// TIA Portal V19 export
// export: Created 2026-10-15T09:44:23.7628945Z, ExportSetting WithDefaults, DisplayName Totally Integrated Automation Portal, DisplayVersion V19, DisplayName TIA Portal Openness, DisplayVersion V19, DisplayName TIA Portal Version Control Interface, DisplayVersion V19, DisplayName STEP 7 Professional, DisplayVersion V19, DisplayName STEP 7 Safety, DisplayVersion V19, DisplayName WinCC Basic/Comfort/Advanced, DisplayVersion V19, DisplayName WinCC Unified, DisplayVersion V19
FUNCTION "ROLL_PB9" : Void   // FC19, SCL
{ S7_Optimized_Access := 'TRUE' }
VERSION : 0.1
// stored: AutoNumber true, IsIECCheckEnabled false, SetENOAutomatically false, UDAEnableTagReadback false
   VAR_TEMP
      r : Bool;
      a1 : Word;
      a2 : Word;
      activeDataBlock : Int;
      comparisonResults : Array[0..0] of Bool;
   END_VAR
BEGIN

   #r := FALSE;
   #a1 := W#16#0000;
   #a2 := W#16#0000;
   #activeDataBlock := 0;
   // PB9, STEP 5 network 1
   #r := ((NOT "ROLL_State".M[32, 1]) AND (NOT "ROLL_State".M[32, 2]) AND "ROLL_IO".Input[0, 2]);
   "ROLL_State".M[32, 0] := #r;
   // PB9, STEP 5 network 2
   #r := "ROLL_State".M[32, 0];
   IF #r THEN
       "ROLL_State".M[32, 1] := TRUE;
   END_IF;
   #r := ((NOT "ROLL_IO".Input[0, 2]) OR "ROLL_IO".Input[0, 1] OR "ROLL_State".M[32, 2]);
   IF #r THEN
       "ROLL_State".M[32, 1] := FALSE;
   END_IF;
   // PB9, STEP 5 network 3
   #r := ((NOT "ROLL_IO".Input[0, 2]) OR "ROLL_IO".Input[0, 1]);
   "ROLL_State".M[32, 2] := #r;
   // PB9, STEP 5 network 4
   #r := ((NOT "ROLL_State".M[12, 0]) AND (NOT "ROLL_State".M[5, 0]) AND (NOT "ROLL_State".M[5, 2]) AND (NOT "ROLL_State".M[9, 0]));
   "ROLL_State".M[35, 1] := #r;
   // PB9, STEP 5 network 5
   #r := "ROLL_IO".Input[0, 4];
   IF #r THEN
       "ROLL_State".M[35, 2] := TRUE;
   END_IF;
   #r := ((NOT "ROLL_State".M[29, 0]) OR (NOT "ROLL_State".M[31, 5]) OR (NOT "ROLL_State".M[35, 1]) OR "ROLL_State".M[16, 3]);
   IF #r THEN
       "ROLL_State".M[35, 2] := FALSE;
   END_IF;
   // PB9, STEP 5 network 6
   #r := ("ROLL_State".M[32, 0] OR "ROLL_State".M[53, 6]);
   IF #r THEN
       "ROLL_State".M[37, 0] := TRUE;
   END_IF;
   #r := ("ROLL_State".M[32, 2] OR "ROLL_State".M[37, 1] OR "ROLL_State".M[38, 0] OR "ROLL_State".M[39, 5]);
   IF #r THEN
       "ROLL_State".M[37, 0] := FALSE;
   END_IF;
   // PB9, STEP 5 network 7
   #r := ((NOT "ROLL_IO".Input[123, 5]) AND (NOT "ROLL_IO".Input[123, 6]) AND (NOT "ROLL_State".M[53, 6]) AND "ROLL_State".M[31, 5] AND "ROLL_State".M[35, 2] AND "ROLL_State".M[37, 0]);
   IF #r THEN
       "ROLL_State".M[37, 1] := TRUE;
   END_IF;
   #r := ("ROLL_State".M[32, 2] OR "ROLL_State".M[37, 2] OR "ROLL_State".M[39, 6]);
   IF #r THEN
       "ROLL_State".M[37, 1] := FALSE;
   END_IF;
   // PB9, STEP 5 network 8
   #r := ((NOT "ROLL_IO".Output[113, 3]) AND (NOT "ROLL_State".M[9, 1]) AND (("ROLL_IO".Input[0, 5] AND "ROLL_IO".Input[14, 3] AND "ROLL_State".M[0, 4]) OR ("ROLL_IO".Input[123, 4] AND "ROLL_IO".Input[124, 4] AND "ROLL_State".M[0, 3])) AND "ROLL_State".M[35, 2] AND "ROLL_State".M[37, 1]);
   IF #r THEN
       "ROLL_State".M[37, 2] := TRUE;
   END_IF;
   #r := ("ROLL_State".M[32, 2] OR "ROLL_State".M[37, 3]);
   IF #r THEN
       "ROLL_State".M[37, 2] := FALSE;
   END_IF;
   // PB9, STEP 5 network 9
   #r := ((NOT "ROLL_State".M[16, 0]) AND (NOT "ROLL_State".M[16, 1]) AND (NOT "ROLL_State".M[16, 4]) AND (NOT "ROLL_State".M[191, 5]) AND "ROLL_IO".Input[14, 0] AND "ROLL_State".M[190, 1] AND "ROLL_State".M[191, 4] AND "ROLL_State".M[35, 2] AND "ROLL_State".M[37, 2]);
   IF #r THEN
       "ROLL_State".M[37, 3] := TRUE;
   END_IF;
   #r := ("ROLL_State".M[32, 2] OR "ROLL_State".M[37, 5] OR "ROLL_State".M[40, 0]);
   IF #r THEN
       "ROLL_State".M[37, 3] := FALSE;
   END_IF;
   // PB9, STEP 5 network 10
   #r := ((NOT "ROLL_IO".Input[123, 5]) AND (NOT "ROLL_IO".Input[123, 6]) AND "ROLL_IO".Input[124, 1] AND "ROLL_IO".Input[124, 4] AND "ROLL_State".M[0, 3] AND "ROLL_State".M[35, 2] AND "ROLL_State".M[37, 3]);
   IF #r THEN
       "ROLL_State".M[37, 5] := TRUE;
   END_IF;
   #r := ("ROLL_State".M[32, 2] OR "ROLL_State".M[37, 6]);
   IF #r THEN
       "ROLL_State".M[37, 5] := FALSE;
   END_IF;
   // PB9, STEP 5 network 11
   #r := ((NOT "ROLL_IO".Output[113, 2]) AND "ROLL_IO".Output[113, 3] AND "ROLL_State".M[35, 2] AND "ROLL_State".M[37, 5] AND "ROLL_State".S5Timers[18].Q);
   IF #r THEN
       "ROLL_State".M[37, 6] := TRUE;
   END_IF;
   #r := ("ROLL_State".M[32, 2] OR "ROLL_State".M[37, 7]);
   IF #r THEN
       "ROLL_State".M[37, 6] := FALSE;
   END_IF;
   // PB9, STEP 5 network 12
   #r := ((NOT "ROLL_State".M[37, 5]) AND "ROLL_State".M[35, 2] AND "ROLL_State".M[37, 6]);
   IF #r THEN
       "ROLL_State".M[37, 7] := TRUE;
   END_IF;
   #r := ("ROLL_State".M[32, 2] OR "ROLL_State".M[38, 0]);
   IF #r THEN
       "ROLL_State".M[37, 7] := FALSE;
   END_IF;
   // PB9, STEP 5 network 13
   #r := ((NOT "ROLL_State".M[70, 2]) AND (((NOT "ROLL_IO".Output[113, 2]) AND "ROLL_IO".Output[113, 3] AND "ROLL_IO".Input[124, 4] AND "ROLL_State".M[28, 4] AND "ROLL_State".M[37, 0]) OR ("ROLL_State".M[37, 7] AND "ROLL_State".S5Timers[20].Q)) AND "ROLL_IO".Input[123, 5] AND "ROLL_State".M[35, 2]);
   IF #r THEN
       "ROLL_State".M[38, 0] := TRUE;
   END_IF;
   #r := ("ROLL_State".M[32, 2] OR "ROLL_State".M[39, 4]);
   IF #r THEN
       "ROLL_State".M[38, 0] := FALSE;
   END_IF;
   // PB9, STEP 5 network 14
   #r := ((NOT "ROLL_IO".Input[124, 5]) AND "ROLL_IO".Input[124, 4] AND "ROLL_State".M[35, 2] AND "ROLL_State".M[38, 0]);
   IF #r THEN
       "ROLL_State".M[39, 4] := TRUE;
   END_IF;
   #r := ("ROLL_State".M[32, 2] OR "ROLL_State".M[39, 5]);
   IF #r THEN
       "ROLL_State".M[39, 4] := FALSE;
   END_IF;
   // PB9, STEP 5 network 15
   #r := ((NOT "ROLL_IO".Input[124, 4]) AND (("ROLL_State".M[28, 4] AND "ROLL_State".M[37, 0]) OR "ROLL_State".M[39, 4]) AND "ROLL_IO".Input[124, 5] AND "ROLL_State".M[35, 2]);
   IF #r THEN
       "ROLL_State".M[39, 5] := TRUE;
   END_IF;
   #r := ("ROLL_State".M[32, 2] OR "ROLL_State".M[39, 6]);
   IF #r THEN
       "ROLL_State".M[39, 5] := FALSE;
   END_IF;
   // PB9, STEP 5 network 16
   #r := ((NOT "ROLL_IO".Input[124, 2]) AND "ROLL_IO".Input[11, 0] AND "ROLL_IO".Input[11, 6] AND "ROLL_IO".Input[12, 1] AND "ROLL_IO".Input[12, 7] AND "ROLL_IO".Input[124, 1] AND "ROLL_State".M[35, 2] AND "ROLL_State".M[39, 5]);
   IF #r THEN
       "ROLL_State".M[39, 6] := TRUE;
   END_IF;
   #r := ("ROLL_State".M[32, 2] OR "ROLL_State".M[39, 7]);
   IF #r THEN
       "ROLL_State".M[39, 6] := FALSE;
   END_IF;
   // PB9, STEP 5 network 17
   #r := ((NOT "ROLL_IO".Input[124, 1]) AND "ROLL_IO".Input[124, 2] AND "ROLL_State".M[35, 2] AND "ROLL_State".M[39, 6]);
   IF #r THEN
       "ROLL_State".M[39, 7] := TRUE;
   END_IF;
   #r := ("ROLL_State".M[32, 2] OR "ROLL_State".M[40, 0]);
   IF #r THEN
       "ROLL_State".M[39, 7] := FALSE;
   END_IF;
   // PB9, STEP 5 network 18
   #r := ((NOT "ROLL_IO".Input[12, 5]) AND ("ROLL_State".M[37, 3] OR "ROLL_State".M[39, 7]) AND "ROLL_IO".Input[11, 0] AND "ROLL_IO".Input[11, 6] AND "ROLL_IO".Input[12, 1] AND "ROLL_IO".Input[12, 7] AND "ROLL_State".M[35, 2]);
   IF #r THEN
       "ROLL_State".M[40, 0] := TRUE;
   END_IF;
   #r := ("ROLL_State".M[32, 2] OR "ROLL_State".M[40, 1]);
   IF #r THEN
       "ROLL_State".M[40, 0] := FALSE;
   END_IF;
   // PB9, STEP 5 network 19
   #r := ("ROLL_IO".Input[12, 5] AND "ROLL_IO".Input[12, 7] AND "ROLL_State".M[35, 2] AND "ROLL_State".M[40, 0]);
   IF #r THEN
       "ROLL_State".M[40, 1] := TRUE;
   END_IF;
   #r := ("ROLL_State".M[32, 2] OR "ROLL_State".M[40, 2] OR "ROLL_State".M[41, 6] OR "ROLL_State".M[43, 2] OR "ROLL_State".M[44, 7] OR "ROLL_State".M[46, 2] OR "ROLL_State".M[47, 6] OR "ROLL_State".M[49, 2] OR "ROLL_State".M[50, 6]);
   IF #r THEN
       "ROLL_State".M[40, 1] := FALSE;
   END_IF;
   // PB9, STEP 5 network 20
   #r := ((NOT "ROLL_IO".Input[11, 1]) AND "ROLL_IO".Input[11, 0] AND "ROLL_State".M[110, 0] AND "ROLL_State".M[35, 2] AND "ROLL_State".M[40, 1] AND "ROLL_State".M[63, 1]);
   IF #r THEN
       "ROLL_State".M[40, 2] := TRUE;
   END_IF;
   #r := ("ROLL_State".M[32, 2] OR "ROLL_State".M[40, 3]);
   IF #r THEN
       "ROLL_State".M[40, 2] := FALSE;
   END_IF;
   // PB9, STEP 5 network 21
   #r := ("ROLL_IO".Input[11, 1] AND "ROLL_IO".Input[11, 6] AND "ROLL_State".M[35, 2] AND "ROLL_State".M[40, 2]);
   IF #r THEN
       "ROLL_State".M[40, 3] := TRUE;
   END_IF;
   #r := ("ROLL_State".M[32, 2] OR "ROLL_State".M[40, 4]);
   IF #r THEN
       "ROLL_State".M[40, 3] := FALSE;
   END_IF;
   // PB9, STEP 5 network 22
   #r := ((NOT "ROLL_IO".Input[12, 1]) AND "ROLL_IO".Input[12, 5] AND "ROLL_State".M[35, 2] AND "ROLL_State".M[40, 3]);
   IF #r THEN
       "ROLL_State".M[40, 4] := TRUE;
   END_IF;
   #r := ("ROLL_State".M[32, 2] OR "ROLL_State".M[40, 5]);
   IF #r THEN
       "ROLL_State".M[40, 4] := FALSE;
   END_IF;
   // PB9, STEP 5 network 23
   #r := ("ROLL_IO".Input[12, 1] AND "ROLL_IO".Input[12, 7] AND "ROLL_State".M[35, 2] AND "ROLL_State".M[40, 4]);
   IF #r THEN
       "ROLL_State".M[40, 5] := TRUE;
   END_IF;
   #r := ("ROLL_State".M[32, 2] OR "ROLL_State".M[40, 6]);
   IF #r THEN
       "ROLL_State".M[40, 5] := FALSE;
   END_IF;
   // PB9, STEP 5 network 24
   #r := ("ROLL_State".M[35, 2] AND "ROLL_State".M[40, 5] AND "ROLL_State".S5Timers[1].Q);
   IF #r THEN
       "ROLL_State".M[40, 6] := TRUE;
   END_IF;
   #r := ("ROLL_State".M[32, 2] OR "ROLL_State".M[40, 7]);
   IF #r THEN
       "ROLL_State".M[40, 6] := FALSE;
   END_IF;
   // PB9, STEP 5 network 25
   #r := ("ROLL_State".M[35, 2] AND "ROLL_State".M[40, 6]);
   IF #r THEN
       "ROLL_State".M[40, 7] := TRUE;
   END_IF;
   #r := ("ROLL_State".M[32, 2] OR "ROLL_State".M[41, 0]);
   IF #r THEN
       "ROLL_State".M[40, 7] := FALSE;
   END_IF;
   // PB9, STEP 5 network 26
   #r := ((NOT "ROLL_IO".Input[12, 5]) AND (("ROLL_IO".Input[13, 3] AND "ROLL_State".M[63, 1]) OR (NOT "ROLL_State".M[111, 5])) AND "ROLL_State".M[35, 2] AND "ROLL_State".M[40, 7]);
   IF #r THEN
       "ROLL_State".M[41, 0] := TRUE;
   END_IF;
   #r := ("ROLL_State".M[32, 2] OR "ROLL_State".M[41, 1]);
   IF #r THEN
       "ROLL_State".M[41, 0] := FALSE;
   END_IF;
   // PB9, STEP 5 network 27
   #r := ("ROLL_IO".Input[12, 5] AND "ROLL_IO".Input[12, 7] AND "ROLL_State".M[35, 2] AND "ROLL_State".M[41, 0]);
   IF #r THEN
       "ROLL_State".M[41, 1] := TRUE;
   END_IF;
   #r := ("ROLL_State".M[32, 2] OR "ROLL_State".M[41, 2]);
   IF #r THEN
       "ROLL_State".M[41, 1] := FALSE;
   END_IF;
   // PB9, STEP 5 network 28
   #r := ("ROLL_State".M[35, 2] AND "ROLL_State".M[41, 1] AND "ROLL_State".S5Timers[2].Q);
   IF #r THEN
       "ROLL_State".M[41, 2] := TRUE;
   END_IF;
   #r := ("ROLL_State".M[32, 2] OR "ROLL_State".M[41, 3] OR "ROLL_State".M[41, 6] OR "ROLL_State".M[43, 2] OR "ROLL_State".M[44, 7] OR "ROLL_State".M[46, 2] OR "ROLL_State".M[47, 6] OR "ROLL_State".M[49, 2]);
   IF #r THEN
       "ROLL_State".M[41, 2] := FALSE;
   END_IF;
   // PB9, STEP 5 network 29
   #r := ((NOT "ROLL_State".M[110, 1]) AND (NOT "ROLL_State".M[110, 2]) AND "ROLL_State".M[35, 2] AND "ROLL_State".M[41, 2]);
   IF #r THEN
       "ROLL_State".M[41, 3] := TRUE;
   END_IF;
   #r := ("ROLL_State".M[32, 2] OR "ROLL_State".M[41, 4]);
   IF #r THEN
       "ROLL_State".M[41, 3] := FALSE;
   END_IF;
   // PB9, STEP 5 network 30
   #r := ("ROLL_IO".Input[13, 3] AND "ROLL_State".M[35, 2] AND "ROLL_State".M[41, 3] AND "ROLL_State".M[63, 1]);
   IF #r THEN
       "ROLL_State".M[41, 4] := TRUE;
   END_IF;
   #r := ("ROLL_State".M[32, 2] OR "ROLL_State".M[44, 7] OR "ROLL_State".M[50, 6] OR "ROLL_State".M[52, 0]);
   IF #r THEN
       "ROLL_State".M[41, 4] := FALSE;
   END_IF;
   // PB9, STEP 5 network 31
   #r := ((NOT "ROLL_IO".Input[11, 2]) AND (((NOT "ROLL_State".M[110, 0]) AND "ROLL_State".M[40, 1]) OR "ROLL_State".M[41, 2]) AND "ROLL_IO".Input[12, 5] AND "ROLL_IO".Input[12, 7] AND "ROLL_State".M[110, 1] AND "ROLL_State".M[35, 2]);
   IF #r THEN
       "ROLL_State".M[41, 6] := TRUE;
   END_IF;
   #r := ("ROLL_State".M[32, 2] OR "ROLL_State".M[41, 7]);
   IF #r THEN
       "ROLL_State".M[41, 6] := FALSE;
   END_IF;
   // PB9, STEP 5 network 32
   #r := ("ROLL_IO".Input[11, 2] AND "ROLL_IO".Input[11, 6] AND "ROLL_State".M[35, 2] AND "ROLL_State".M[41, 6]);
   IF #r THEN
       "ROLL_State".M[41, 7] := TRUE;
   END_IF;
   #r := ("ROLL_State".M[32, 2] OR "ROLL_State".M[42, 0]);
   IF #r THEN
       "ROLL_State".M[41, 7] := FALSE;
   END_IF;
   // PB9, STEP 5 network 33
   #r := ((NOT "ROLL_IO".Input[12, 1]) AND "ROLL_IO".Input[12, 5] AND "ROLL_State".M[35, 2] AND "ROLL_State".M[41, 7]);
   IF #r THEN
       "ROLL_State".M[42, 0] := TRUE;
   END_IF;
   #r := ("ROLL_State".M[32, 2] OR "ROLL_State".M[42, 1]);
   IF #r THEN
       "ROLL_State".M[42, 0] := FALSE;
   END_IF;
   // PB9, STEP 5 network 34
   #r := ("ROLL_IO".Input[12, 1] AND "ROLL_IO".Input[12, 7] AND "ROLL_State".M[35, 2] AND "ROLL_State".M[42, 0]);
   IF #r THEN
       "ROLL_State".M[42, 1] := TRUE;
   END_IF;
   #r := ("ROLL_State".M[32, 2] OR "ROLL_State".M[42, 2]);
   IF #r THEN
       "ROLL_State".M[42, 1] := FALSE;
   END_IF;
   // PB9, STEP 5 network 35
   #r := ("ROLL_State".M[35, 2] AND "ROLL_State".M[42, 1] AND "ROLL_State".S5Timers[1].Q);
   IF #r THEN
       "ROLL_State".M[42, 2] := TRUE;
   END_IF;
   #r := ("ROLL_State".M[32, 2] OR "ROLL_State".M[42, 3]);
   IF #r THEN
       "ROLL_State".M[42, 2] := FALSE;
   END_IF;
   // PB9, STEP 5 network 36
   #r := ("ROLL_State".M[35, 2] AND "ROLL_State".M[42, 2]);
   IF #r THEN
       "ROLL_State".M[42, 3] := TRUE;
   END_IF;
   #r := ("ROLL_State".M[32, 2] OR "ROLL_State".M[42, 4]);
   IF #r THEN
       "ROLL_State".M[42, 3] := FALSE;
   END_IF;
   // PB9, STEP 5 network 37
   #r := ((NOT "ROLL_IO".Input[12, 5]) AND (("ROLL_IO".Input[13, 3] AND "ROLL_State".M[63, 1]) OR (NOT "ROLL_State".M[111, 5])) AND "ROLL_State".M[35, 2] AND "ROLL_State".M[42, 3]);
   IF #r THEN
       "ROLL_State".M[42, 4] := TRUE;
   END_IF;
   #r := ("ROLL_State".M[32, 2] OR "ROLL_State".M[42, 5]);
   IF #r THEN
       "ROLL_State".M[42, 4] := FALSE;
   END_IF;
   // PB9, STEP 5 network 38
   #r := ("ROLL_IO".Input[12, 5] AND "ROLL_IO".Input[12, 7] AND "ROLL_State".M[35, 2] AND "ROLL_State".M[42, 4]);
   IF #r THEN
       "ROLL_State".M[42, 5] := TRUE;
   END_IF;
   #r := ("ROLL_State".M[32, 2] OR "ROLL_State".M[42, 6]);
   IF #r THEN
       "ROLL_State".M[42, 5] := FALSE;
   END_IF;
   // PB9, STEP 5 network 39
   #r := ("ROLL_State".M[35, 2] AND "ROLL_State".M[42, 5] AND "ROLL_State".S5Timers[2].Q);
   IF #r THEN
       "ROLL_State".M[42, 6] := TRUE;
   END_IF;
   #r := ("ROLL_State".M[32, 2] OR "ROLL_State".M[42, 7] OR "ROLL_State".M[43, 2] OR "ROLL_State".M[44, 7] OR "ROLL_State".M[46, 2] OR "ROLL_State".M[47, 6] OR "ROLL_State".M[49, 2]);
   IF #r THEN
       "ROLL_State".M[42, 6] := FALSE;
   END_IF;
   // PB9, STEP 5 network 40
   #r := ((NOT "ROLL_State".M[110, 2]) AND "ROLL_State".M[35, 2] AND "ROLL_State".M[42, 6]);
   IF #r THEN
       "ROLL_State".M[42, 7] := TRUE;
   END_IF;
   #r := ("ROLL_State".M[32, 2] OR "ROLL_State".M[43, 0]);
   IF #r THEN
       "ROLL_State".M[42, 7] := FALSE;
   END_IF;
   // PB9, STEP 5 network 41
   #r := ("ROLL_IO".Input[13, 3] AND "ROLL_State".M[35, 2] AND "ROLL_State".M[42, 7] AND "ROLL_State".M[63, 1]);
   IF #r THEN
       "ROLL_State".M[43, 0] := TRUE;
   END_IF;
   #r := ("ROLL_State".M[32, 2] OR "ROLL_State".M[44, 7] OR "ROLL_State".M[50, 6] OR "ROLL_State".M[52, 0]);
   IF #r THEN
       "ROLL_State".M[43, 0] := FALSE;
   END_IF;
   // PB9, STEP 5 network 42
   #r := ((NOT "ROLL_IO".Input[11, 3]) AND (((NOT "ROLL_State".M[110, 0]) AND (NOT "ROLL_State".M[110, 1]) AND "ROLL_State".M[40, 1]) OR ((NOT "ROLL_State".M[110, 1]) AND "ROLL_State".M[41, 2]) OR "ROLL_State".M[42, 6]) AND "ROLL_IO".Input[12, 5] AND "ROLL_IO".Input[12, 7] AND "ROLL_State".M[110, 2] AND "ROLL_State".M[35, 2]);
   IF #r THEN
       "ROLL_State".M[43, 2] := TRUE;
   END_IF;
   #r := ("ROLL_State".M[32, 2] OR "ROLL_State".M[43, 3]);
   IF #r THEN
       "ROLL_State".M[43, 2] := FALSE;
   END_IF;
   // PB9, STEP 5 network 43
   #r := ("ROLL_IO".Input[11, 3] AND "ROLL_IO".Input[11, 6] AND "ROLL_State".M[35, 2] AND "ROLL_State".M[43, 2]);
   IF #r THEN
       "ROLL_State".M[43, 3] := TRUE;
   END_IF;
   #r := ("ROLL_State".M[32, 2] OR "ROLL_State".M[43, 4]);
   IF #r THEN
       "ROLL_State".M[43, 3] := FALSE;
   END_IF;
   // PB9, STEP 5 network 44
   #r := ((NOT "ROLL_IO".Input[12, 1]) AND "ROLL_IO".Input[12, 5] AND "ROLL_State".M[35, 2] AND "ROLL_State".M[43, 3]);
   IF #r THEN
       "ROLL_State".M[43, 4] := TRUE;
   END_IF;
   #r := ("ROLL_State".M[32, 2] OR "ROLL_State".M[43, 5]);
   IF #r THEN
       "ROLL_State".M[43, 4] := FALSE;
   END_IF;
   // PB9, STEP 5 network 45
   #r := ("ROLL_IO".Input[12, 1] AND "ROLL_IO".Input[12, 7] AND "ROLL_State".M[35, 2] AND "ROLL_State".M[43, 4]);
   IF #r THEN
       "ROLL_State".M[43, 5] := TRUE;
   END_IF;
   #r := ("ROLL_State".M[32, 2] OR "ROLL_State".M[43, 6]);
   IF #r THEN
       "ROLL_State".M[43, 5] := FALSE;
   END_IF;
   // PB9, STEP 5 network 46
   #r := ("ROLL_State".M[35, 2] AND "ROLL_State".M[43, 5] AND "ROLL_State".S5Timers[1].Q);
   IF #r THEN
       "ROLL_State".M[43, 6] := TRUE;
   END_IF;
   #r := ("ROLL_State".M[32, 2] OR "ROLL_State".M[43, 7]);
   IF #r THEN
       "ROLL_State".M[43, 6] := FALSE;
   END_IF;
   // PB9, STEP 5 network 47
   #r := ("ROLL_State".M[35, 2] AND "ROLL_State".M[43, 6]);
   IF #r THEN
       "ROLL_State".M[43, 7] := TRUE;
   END_IF;
   #r := ("ROLL_State".M[32, 2] OR "ROLL_State".M[44, 0]);
   IF #r THEN
       "ROLL_State".M[43, 7] := FALSE;
   END_IF;
   // PB9, STEP 5 network 48
   #r := ((NOT "ROLL_IO".Input[12, 5]) AND (("ROLL_IO".Input[13, 3] AND "ROLL_State".M[63, 1]) OR (NOT "ROLL_State".M[111, 5])) AND "ROLL_State".M[35, 2] AND "ROLL_State".M[43, 7]);
   IF #r THEN
       "ROLL_State".M[44, 0] := TRUE;
   END_IF;
   #r := ("ROLL_State".M[32, 2] OR "ROLL_State".M[44, 1]);
   IF #r THEN
       "ROLL_State".M[44, 0] := FALSE;
   END_IF;
   // PB9, STEP 5 network 49
   #r := ("ROLL_IO".Input[12, 5] AND "ROLL_IO".Input[12, 7] AND "ROLL_State".M[35, 2] AND "ROLL_State".M[44, 0]);
   IF #r THEN
       "ROLL_State".M[44, 1] := TRUE;
   END_IF;
   #r := ("ROLL_State".M[32, 2] OR "ROLL_State".M[44, 2]);
   IF #r THEN
       "ROLL_State".M[44, 1] := FALSE;
   END_IF;
   // PB9, STEP 5 network 50
   #r := ("ROLL_State".M[35, 2] AND "ROLL_State".M[44, 1] AND "ROLL_State".S5Timers[2].Q);
   IF #r THEN
       "ROLL_State".M[44, 2] := TRUE;
   END_IF;
   #r := ("ROLL_State".M[32, 2] OR "ROLL_State".M[44, 3] OR "ROLL_State".M[44, 7] OR "ROLL_State".M[46, 2] OR "ROLL_State".M[47, 6] OR "ROLL_State".M[49, 2]);
   IF #r THEN
       "ROLL_State".M[44, 2] := FALSE;
   END_IF;
   // PB9, STEP 5 network 51
   #r := ("ROLL_State".M[35, 2] AND "ROLL_State".M[44, 2]);
   IF #r THEN
       "ROLL_State".M[44, 3] := TRUE;
   END_IF;
   #r := ("ROLL_State".M[32, 2] OR "ROLL_State".M[44, 4]);
   IF #r THEN
       "ROLL_State".M[44, 3] := FALSE;
   END_IF;
   // PB9, STEP 5 network 52
   #r := ("ROLL_IO".Input[13, 3] AND "ROLL_State".M[35, 2] AND "ROLL_State".M[44, 3] AND "ROLL_State".M[63, 1]);
   IF #r THEN
       "ROLL_State".M[44, 4] := TRUE;
   END_IF;
   #r := ("ROLL_State".M[32, 2] OR "ROLL_State".M[44, 7] OR "ROLL_State".M[50, 6] OR "ROLL_State".M[52, 0]);
   IF #r THEN
       "ROLL_State".M[44, 4] := FALSE;
   END_IF;
   // PB9, STEP 5 network 53
   #r := (((NOT "ROLL_State".M[110, 0]) AND (NOT "ROLL_State".M[110, 1]) AND (NOT "ROLL_State".M[110, 2]) AND "ROLL_State".M[40, 1]) OR ((NOT "ROLL_State".M[110, 1]) AND (NOT "ROLL_State".M[110, 2]) AND "ROLL_State".M[41, 4]) OR ((NOT "ROLL_State".M[110, 2]) AND "ROLL_State".M[43, 0]) OR "ROLL_State".M[44, 4]);
   "ROLL_State".M[240, 0] := #r;
   // PB9, STEP 5 network 54
   #r := ((NOT "ROLL_IO".Input[11, 4]) AND "ROLL_IO".Input[12, 5] AND "ROLL_IO".Input[12, 7] AND "ROLL_State".M[110, 3] AND "ROLL_State".M[240, 0] AND "ROLL_State".M[35, 2] AND "ROLL_State".M[63, 1]);
   IF #r THEN
       "ROLL_State".M[44, 7] := TRUE;
   END_IF;
   #r := ("ROLL_State".M[32, 2] OR "ROLL_State".M[45, 0]);
   IF #r THEN
       "ROLL_State".M[44, 7] := FALSE;
   END_IF;
   // PB9, STEP 5 network 55
   #r := ("ROLL_IO".Input[11, 4] AND "ROLL_IO".Input[11, 6] AND "ROLL_State".M[35, 2] AND "ROLL_State".M[44, 7]);
   IF #r THEN
       "ROLL_State".M[45, 0] := TRUE;
   END_IF;
   #r := ("ROLL_State".M[32, 2] OR "ROLL_State".M[45, 1]);
   IF #r THEN
       "ROLL_State".M[45, 0] := FALSE;
   END_IF;
   // PB9, STEP 5 network 56
   #r := ((NOT "ROLL_IO".Input[12, 1]) AND "ROLL_IO".Input[12, 5] AND "ROLL_State".M[35, 2] AND "ROLL_State".M[45, 0]);
   IF #r THEN
       "ROLL_State".M[45, 1] := TRUE;
   END_IF;
   #r := ("ROLL_State".M[32, 2] OR "ROLL_State".M[45, 2]);
   IF #r THEN
       "ROLL_State".M[45, 1] := FALSE;
   END_IF;
   // PB9, STEP 5 network 57
   #r := ("ROLL_IO".Input[12, 1] AND "ROLL_IO".Input[12, 7] AND "ROLL_State".M[35, 2] AND "ROLL_State".M[45, 1]);
   IF #r THEN
       "ROLL_State".M[45, 2] := TRUE;
   END_IF;
   #r := ("ROLL_State".M[32, 2] OR "ROLL_State".M[45, 3]);
   IF #r THEN
       "ROLL_State".M[45, 2] := FALSE;
   END_IF;
   // PB9, STEP 5 network 58
   #r := ("ROLL_State".M[35, 2] AND "ROLL_State".M[45, 2] AND "ROLL_State".S5Timers[1].Q);
   IF #r THEN
       "ROLL_State".M[45, 3] := TRUE;
   END_IF;
   #r := ("ROLL_State".M[32, 2] OR "ROLL_State".M[45, 4]);
   IF #r THEN
       "ROLL_State".M[45, 3] := FALSE;
   END_IF;
   // PB9, STEP 5 network 59
   #r := ("ROLL_State".M[35, 2] AND "ROLL_State".M[45, 3]);
   IF #r THEN
       "ROLL_State".M[45, 4] := TRUE;
   END_IF;
   #r := ("ROLL_State".M[32, 2] OR "ROLL_State".M[45, 5]);
   IF #r THEN
       "ROLL_State".M[45, 4] := FALSE;
   END_IF;
   // PB9, STEP 5 network 60
   #r := ((NOT "ROLL_IO".Input[12, 5]) AND "ROLL_State".M[35, 2] AND "ROLL_State".M[45, 4]);
   IF #r THEN
       "ROLL_State".M[45, 5] := TRUE;
   END_IF;
   #r := ("ROLL_State".M[32, 2] OR "ROLL_State".M[45, 6]);
   IF #r THEN
       "ROLL_State".M[45, 5] := FALSE;
   END_IF;
   // PB9, STEP 5 network 61
   #r := ("ROLL_IO".Input[12, 5] AND "ROLL_IO".Input[12, 7] AND "ROLL_State".M[35, 2] AND "ROLL_State".M[45, 5]);
   IF #r THEN
       "ROLL_State".M[45, 6] := TRUE;
   END_IF;
   #r := ("ROLL_State".M[32, 2] OR "ROLL_State".M[45, 7]);
   IF #r THEN
       "ROLL_State".M[45, 6] := FALSE;
   END_IF;
   // PB9, STEP 5 network 62
   #r := (("ROLL_State".M[0, 4] OR "ROLL_State".S5Timers[2].Q) AND "ROLL_State".M[35, 2] AND "ROLL_State".M[45, 6]);
   IF #r THEN
       "ROLL_State".M[45, 7] := TRUE;
   END_IF;
   #r := ("ROLL_State".M[32, 2] OR "ROLL_State".M[46, 0] OR "ROLL_State".M[46, 2] OR "ROLL_State".M[47, 6] OR "ROLL_State".M[49, 2]);
   IF #r THEN
       "ROLL_State".M[45, 7] := FALSE;
   END_IF;
   // PB9, STEP 5 network 63
   #r := ("ROLL_State".M[35, 2] AND "ROLL_State".M[45, 7]);
   IF #r THEN
       "ROLL_State".M[46, 0] := TRUE;
   END_IF;
   #r := ("ROLL_State".M[32, 2] OR "ROLL_State".M[46, 1]);
   IF #r THEN
       "ROLL_State".M[46, 0] := FALSE;
   END_IF;
   // PB9, STEP 5 network 64
   #r := ("ROLL_IO".Input[13, 3] AND "ROLL_State".M[35, 2] AND "ROLL_State".M[46, 0] AND "ROLL_State".M[63, 1]);
   IF #r THEN
       "ROLL_State".M[46, 1] := TRUE;
   END_IF;
   #r := ("ROLL_State".M[32, 2] OR "ROLL_State".M[50, 6] OR "ROLL_State".M[52, 0]);
   IF #r THEN
       "ROLL_State".M[46, 1] := FALSE;
   END_IF;
   // PB9, STEP 5 network 65
   RETURN;
END_FUNCTION
